FUNCTION_BLOCK TransportHandlingCAT (* CAT Function Block Type *)
  (* Standard: 61499-2 *)
  (* Version 0.0, 7/7/2026, template *)
  PACKAGE Main;
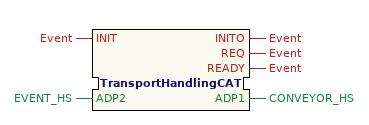
  EVENT_INPUT
    INIT; (* Initialization Request *)
  END_EVENT
  EVENT_OUTPUT
    INITO; (* Initialization Confirm *)
    REQ; (* Execution Confirmation *)
    READY;
  END_EVENT
  SOCKETS
    ADP2 : EVENT_HS;
  END_SOCKETS
  PLUGS
    ADP1 : CONVEYOR_HS;
  END_PLUGS
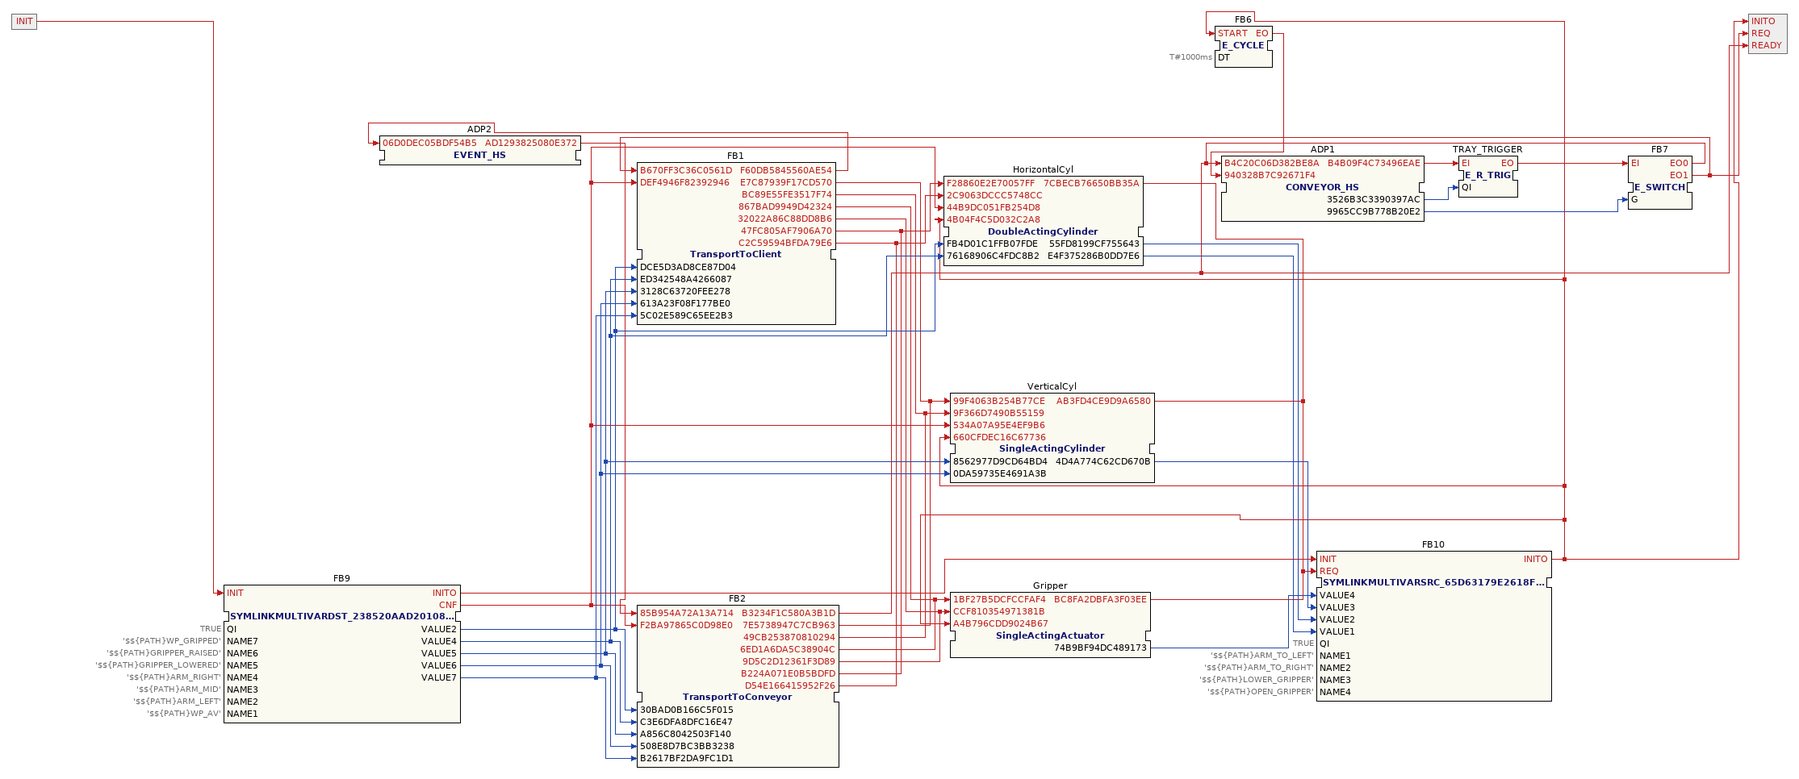
  FBS
    FB1 : TransportToClient;
    FB2 : TransportToConveyor;
    Gripper : SingleActingActuator;
    VerticalCyl : SingleActingCylinder;
    FB6 : E_CYCLE(DT := T#1000ms);
    FB7 : E_SWITCH;
    TRAY_TRIGGER : E_R_TRIG;
    FB9 : SYMLINKMULTIVARDST_238520AAD20108C65(QI := TRUE, NAME7 := '$${PATH}WP_GRIPPED', NAME6 := '$${PATH}GRIPPER_RAISED', NAME5 := '$${PATH}GRIPPER_LOWERED', NAME4 := '$${PATH}ARM_RIGHT', NAME3 := '$${PATH}ARM_MID', NAME2 := '$${PATH}ARM_LEFT', NAME1 := '$${PATH}WP_AV'); {SET_ATTRIBUTE(Configuration.GenericFBType.InterfaceParams, Runtime.System#I:=7;VALUE${I$}:BOOL,BOOL,BOOL,BOOL,BOOL,BOOL,BOOL)}
    FB10 : SYMLINKMULTIVARSRC_65D63179E2618F5E(QI := TRUE, NAME1 := '$${PATH}ARM_TO_LEFT', NAME2 := '$${PATH}ARM_TO_RIGHT', NAME3 := '$${PATH}LOWER_GRIPPER', NAME4 := '$${PATH}OPEN_GRIPPER'); {SET_ATTRIBUTE(Configuration.GenericFBType.InterfaceParams, Runtime.System#I:=5;VALUE${I$}:BOOL,BOOL,BOOL,BOOL,BOOL)}
    HorizontalCyl : DoubleActingCylinder;
  END_FBS
  EVENT_CONNECTIONS
    INIT TO FB9.INIT;
    FB9.INITO TO FB10.INIT;
    ADP2.AD1293825080E372 TO FB2.85B954A72A13A714;
    FB1.F60DB5845560AE54 TO ADP2.06D0DEC05BDF54B5;
    FB1.E7C87939F17CD570 TO VerticalCyl.99F4063B254B77CE;
    FB1.BC89E55FE3517F74 TO VerticalCyl.9F366D7490B55159;
    FB1.867BAD9949D42324 TO Gripper.1BF27B5DCFCCFAF4;
    FB1.32022A86C88DD8B6 TO Gripper.CCF810354971381B;
    FB1.47FC805AF7906A70 TO HorizontalCyl.F28860E2E70057FF;
    FB1.C2C59594BFDA79E6 TO HorizontalCyl.2C9063DCCC5748CC;
    FB2.B3234F1C580A3B1D TO ADP1.B4C20C06D382BE8A;
    FB2.B3234F1C580A3B1D TO READY;
    FB2.7E5738947C7CB963 TO VerticalCyl.99F4063B254B77CE;
    FB2.49CB253870810294 TO VerticalCyl.9F366D7490B55159;
    FB2.6ED1A6DA5C38904C TO Gripper.1BF27B5DCFCCFAF4;
    FB2.9D5C2D12361F3D89 TO Gripper.CCF810354971381B;
    FB2.B224A071E0B5BDFD TO HorizontalCyl.F28860E2E70057FF;
    FB2.D54E166415952F26 TO HorizontalCyl.2C9063DCCC5748CC;
    FB10.INITO TO INITO;
    FB10.INITO TO FB6.START;
    FB6.EO TO ADP1.940328B7C92671F4;
    FB7.EO0 TO ADP1.B4C20C06D382BE8A;
    ADP1.B4B09F4C73496EAE TO TRAY_TRIGGER.EI;
    TRAY_TRIGGER.EO TO FB7.EI;
    FB7.EO1 TO REQ;
    FB7.EO1 TO FB1.B670FF3C36C0561D;
    FB9.CNF TO FB1.DEF4946F82392946;
    FB9.CNF TO FB2.F2BA97865C0D98E0;
    FB9.CNF TO HorizontalCyl.44B9DC051FB254D8;
    FB9.CNF TO VerticalCyl.534A07A95E4EF9B6;
    VerticalCyl.AB3FD4CE9D9A6580 TO FB10.REQ;
    Gripper.BC8FA2DBFA3F03EE TO FB10.REQ;
    HorizontalCyl.7CBECB76650BB35A TO FB10.REQ;
    FB10.INITO TO HorizontalCyl.4B04F4C5D032C2A8;
    FB10.INITO TO VerticalCyl.660CFDEC16C67736;
    FB10.INITO TO Gripper.A4B796CDD9024B67;
  END_CONNECTIONS
  DATA_CONNECTIONS
    FB9.VALUE2 TO FB1.DCE5D3AD8CE87D04;
    FB9.VALUE2 TO FB2.30BAD0B166C5F015;
    FB9.VALUE4 TO FB2.C3E6DFA8DFC16E47;
    FB9.VALUE4 TO FB1.ED342548A4266087;
    FB9.VALUE2 TO HorizontalCyl.FB4D01C1FFB07FDE;
    FB9.VALUE4 TO HorizontalCyl.76168906C4FDC8B2;
    FB9.VALUE5 TO FB2.A856C8042503F140;
    FB9.VALUE5 TO FB1.3128C63720FEE278;
    FB9.VALUE5 TO VerticalCyl.8562977D9CD64BD4;
    FB9.VALUE6 TO FB1.613A23F08F177BE0;
    FB9.VALUE6 TO FB2.508E8D7BC3BB3238;
    FB9.VALUE6 TO VerticalCyl.0DA59735E4691A3B;
    FB9.VALUE7 TO FB2.B2617BF2DA9FC1D1;
    FB9.VALUE7 TO FB1.5C02E589C65EE2B3;
    Gripper.74B9BF94DC489173 TO FB10.VALUE4;
    VerticalCyl.4D4A774C62CD670B TO FB10.VALUE3;
    HorizontalCyl.55FD8199CF755643 TO FB10.VALUE2;
    HorizontalCyl.E4F375286B0DD7E6 TO FB10.VALUE1;
    ADP1.3526B3C3390397AC TO TRAY_TRIGGER.QI;
    ADP1.9965CC9B778B20E2 TO FB7.G;
  END_CONNECTIONS
END_FUNCTION_BLOCK
